(* IEC 61131-3 sources: kns-port-domestic/upstream/plc-process-lib/src/DUTs/Common, 8 files *)

(* ---- E_CmdResult.dut.st ---- *)
// Назначение: результат обработки команды HMI/SCADA или запроса метода
//             (stSts.stCommon.eCmdResult; каждая обработанная команда увеличивает uiCmdSeq).
// Автор:      kr0nsch
// Версия:     0.1.0
// Документ:   docs/ARCHITECTURE.md, раздел «Общие типы»
{attribute 'qualified_only'}
{attribute 'strict'}
TYPE E_CmdResult :
(
    None                 := 0,   // команд ещё не было
    Accepted             := 1,
    RejectedMode         := 2,   // недопустимо в текущем режиме (пуск в Auto; команды в Local/OOS)
    RejectedInterlock    := 3,   // действует защитная блокировка
    RejectedPermit       := 4,   // нет разрешения (в т. ч. ПЧ не готов)
    RejectedInhibit      := 5,   // пауза после останова, лимит пусков, нет напряжения
    RejectedFault        := 6,   // есть отказ; Reset при неснятой причине; PV негодна (ПИД)
    RejectedState        := 7,   // недопустимо в текущем состоянии (OOS при работающем механизме)
    RejectedNotSupported := 8,   // не поддерживается типом (стоп соленоида, Local у AI)
    RejectedCfg          := 9,   // нет корректной конфигурации
    SubstExpired         := 10   // AI/DI: подмена снята по tSubstMax (событие, а не ответ на команду)
) INT;
END_TYPE

(* ---- E_DeviceMode.dut.st ---- *)
// Назначение: режим работы устройства. Значения 0 нет намеренно: 0 в retain или в регистре
//             Modbus значит «не инициализировано» и трактуется как Manual (санитизация во
//             время работы). Приоритет: OutOfService > Local > Auto/Manual.
// Автор:      kr0nsch
// Версия:     0.1.0
// Документ:   docs/ARCHITECTURE.md, раздел «Общие типы»
{attribute 'qualified_only'}
{attribute 'strict'}
TYPE E_DeviceMode :
(
    Auto         := 1,   // автомат: команды от логики (AI/DI: измерение)
    Manual       := 2,   // ручной дистанционный (AI/DI: подмена значения)
    Local        := 3,   // местный: аппаратный переключатель, ПЛК выходами не управляет
    OutOfService := 4    // выведено из работы
) INT;
END_TYPE

(* ---- E_DeviceType.dut.st ---- *)
// Назначение: тип устройства в stSts.stCommon.eDevType. SCADA по нему выбирает фейсплейт,
//             генератор карты Modbus проверяет, что по адресу блока лежит ожидаемое устройство.
// Автор:      kr0nsch
// Версия:     0.1.0
// Документ:   docs/ARCHITECTURE.md, раздел «Общие типы»
{attribute 'qualified_only'}
{attribute 'strict'}
TYPE E_DeviceType :
(
    None         := 0,   // до первого вызова
    AnalogInput  := 1,
    DigitalInput := 2,
    Motor        := 3,
    MotorVfd     := 4,
    Valve        := 5,
    ControlValve := 6,
    Pid          := 7
) INT;
END_TYPE

(* ---- E_Ne107Status.dut.st ---- *)
// Назначение: диагностический статус по NAMUR NE 107. Значения упорядочены по тяжести,
//             сводный статус — MAX (F_Ne107Worst). Порядок F > C > S > M принят по практике
//             агрегации — сверить с текстом NAMUR NE 107.
// Автор:      kr0nsch
// Версия:     0.1.0
// Документ:   docs/ARCHITECTURE.md, раздел «Общие типы»
{attribute 'qualified_only'}
{attribute 'strict'}
TYPE E_Ne107Status :
(
    Good                := 0,   // норма
    MaintenanceRequired := 1,   // M — требуется обслуживание
    OutOfSpecification  := 2,   // S — вне спецификации
    CheckFunction       := 3,   // C — функциональная проверка (подмена, OOS, конфигурация)
    Failure             := 4    // F — отказ
) INT;
END_TYPE

(* ---- ST_DeviceCmd.dut.st ---- *)
// Назначение: общий заголовок команд HMI/SCADA — первое поле stCommon каждой ST_<Dev>Cmd.
//             Импульсные биты ФБ сбрасывает в том же вызове, маски обнуляет после обработки.
// Автор:      kr0nsch
// Версия:     0.1.0
// Документ:   docs/ARCHITECTURE.md, раздел «Общие типы»
{attribute 'qualified_only'}
TYPE ST_DeviceCmd :
STRUCT
    xSetAuto     : BOOL;   // импульс: в Auto (AI/DI: измерение; выход из OOS)
    xSetManual   : BOOL;   // импульс: в Manual (AI/DI: подмена; выход из OOS)
    xSetOos      : BOOL;   // импульс: вывести из работы
    xReset       : BOOL;   // импульс: сброс зафиксированных отказов + квитирование всех тревог
    xAck         : BOOL;   // импульс: квитировать все тревоги (без сброса отказов)
    wAckReq      : WORD;   // маска: квитировать тревоги слотов (бит i = слот i)
    wShelveReq   : WORD;   // маска: отложить тревоги слотов на stCfg.astAlarm[i].tShelveMax
    wUnshelveReq : WORD;   // маска: вернуть отложенные тревоги
END_STRUCT
END_TYPE

(* ---- ST_DeviceRetain.dut.st ---- *)
// Назначение: энергонезависимые данные устройства. Приложение размещает переменную этого
//             типа в объекте Persistent Variables, по переменной на устройство (st<TAG>Retain).
//             Объявление заморожено целиком, включая имена полей: любое изменение типа
//             переинициализирует persistent-переменную (A-13). Новые данные 1.x — только в
//             элементы audiReserve без переименования. SIZEOF = 36 (Control Win V3, 32 бит).
// Автор:      kr0nsch
// Версия:     0.1.0
// Документ:   docs/ARCHITECTURE.md, раздел «Энергонезависимые данные»
{attribute 'qualified_only'}
TYPE ST_DeviceRetain :
STRUCT
    eRemoteMode      : E_DeviceMode := E_DeviceMode.Manual;   // последний дистанционный режим (Auto/Manual)
    xOutOfService    : BOOL;                     // выведено из работы оператором
    udiOpTime_s      : UDINT;                    // наработка всего, с (двигатель — работа; задвижка — ход)
    udiOpCount       : UDINT;                    // операций всего (двигатель — пуски; арматура — циклы)
    udiOpTimeMaint_s : UDINT;                    // наработка с последнего ТО, с
    udiOpCountMaint  : UDINT;                    // операций с последнего ТО
    audiReserve      : ARRAY[0..3] OF UDINT;     // резерв: новые поля без смены раскладки
END_STRUCT
END_TYPE

(* ---- ST_DeviceSts.dut.st ---- *)
// Назначение: общий заголовок состояния — первое поле stCommon каждой ST_<Dev>Sts.
//             Все 14 полей 16-битные: 28 байт, 14 регистров Modbus подряд. Раскладка
//             нормативна (тест Common_SizeOfSts_MatchesRegisterMap).
// Автор:      kr0nsch
// Версия:     0.1.0
// Документ:   docs/ARCHITECTURE.md, раздел «Общие типы»
{attribute 'qualified_only'}
TYPE ST_DeviceSts :
STRUCT
    wStatus     : WORD;              // биты 0–7 по типу устройства, 8–15 общие (DEV_STS_*)
    wFault      : WORD;              // причины отказа (карта по типу)
    wWarning    : WORD;              // предупреждения (карта по типу)
    wCfgErr     : WORD;              // непройденные проверки Cfg (карта по типу)
    eMode       : E_DeviceMode := E_DeviceMode.Manual;
    eNe107      : E_Ne107Status := E_Ne107Status.CheckFunction;   // до первого вызова — «не проверено»
    eCmdResult  : E_CmdResult := E_CmdResult.None;
    uiCmdSeq    : UINT;              // +1 на каждую обработанную команду (по кругу)
    wAlmActive  : WORD;              // бит i: условие тревоги слота i активно (после задержек)
    wAlmUnack   : WORD;              // бит i: тревога слота i не квитирована
    wAlmShelved : WORD;              // бит i: слот отложен оператором (Shelved, ISA-18.2)
    ePrioUnack  : E_AlarmPriority := E_AlarmPriority.None;   // наивысший приоритет среди неквитированных
    eDevType    : E_DeviceType := E_DeviceType.None;         // тип устройства
    wAlmSuppressed : WORD;           // бит i: слот подавлен логикой (SuppressedByDesign); размер кратен 4 байтам
END_STRUCT
END_TYPE

(* ---- U_RealBits.dut.st ---- *)
// Назначение: доступ к битам REAL — F_IsFinite проверяет экспоненту на NaN и ±Inf без
//             сравнения r = r, результат которого зависит от оптимизатора.
// Автор:      kr0nsch
// Версия:     0.1.0
// Документ:   docs/fb/Functions.md
{attribute 'qualified_only'}
TYPE U_RealBits :
UNION
    rValue  : REAL;    // значение
    dwValue : DWORD;   // те же 32 бита (IEEE 754: знак, 8 бит экспоненты, 23 бита мантиссы)
END_UNION
END_TYPE
